Universal Robots URScript: T001_mock-model-v1_edit_perf_rep1.urscript

def task():
  movej([0, -1.57, 1.57, -1.57, -1.57, 0], a=0.5, v=0.2)
  movel(p[0.3, 0.2, 0.4, 0, 3.14, 0], a=0.3, v=0.1)
end
